// TIA Portal V20 export
Screen "RFIDWrite"  1276x673
  ScreenItem "线_1" at 0,68 size 1363x0  Type=HmiLine
  ScreenItem "符号 IO 域_1" at 451,27 size 475x42  Type=HmiSymbolicIOField
  ScreenItem "permanentareaborderrectangle" at 0,0 size 0x0  Type=HmiRectangle
  ScreenItem "Button_Back" at 2,3 size 90x60  Type=HmiButton
  ScreenItem "txtOverview_3" at 1185,3 size 90x60  Type=HmiTextBox
  ScreenItem "Title_OPMode1_ScreenOverview_X390_Y2" at 439,-2 size 500x30  Type=HmiTextBox
